(*
SPDX-FileCopyrightText: © 2026 Oleksandr Tiutyk <trofimich@gmail.com>
SPDX-License-Identifier: MIT
License: https://opensource.org/license/mit
*)

(*!
<summary>
Beckhoff EL2622: 2-channel relay output terminal (230 V AC / 30 V DC, normally open make contacts).
</summary>
<description>
Process image mapping structure for the EL2622 potential-free relay output terminal.
Each channel switches up to 5 A AC/DC for resistive loads or 2 A AC/DC for inductive loads.
The terminal has two make contacts, not changeover contacts, and does not pass through power contacts.
When used for I/O, link located fields or their containing buffers to the matching selected PDOs.
The record is not a packed wire buffer; compiler padding is not part of the device specification.
Unlinked/default values do not prove valid I/O. The caller evaluates bus/channel validity before use.
Use one owner task per instance and externally synchronize other access; multi-field snapshots are not atomic.
Copies store data without creating hardware links. Keep borrowed field references valid while consumers are bound.
This passive record performs no validation, synchronization, configuration or protocol advancement.
</description>
*)
TYPE EL2622 :
STRUCT
	Ch1 AT %Q* : BOOL;
	Ch2 AT %Q* : BOOL;
END_STRUCT
END_TYPE

(* stored: Version 1.1.0.1, ProductVersion 3.1.4026.20
   DUT EL2622: Id {548de5ea-2158-4842-83a7-9a08f9066951} *)
